Staubli VAL3: insertENDSwitch.pgx

public program insertENDSwitch(string x_sKey, num x_nIndex, bool& x_bToSave)
  local num l_i
begin
  if x_nIndex==0 and progTemp:pProgItem[x_sKey].pProgTemplate[x_nIndex].sTRAJname==""
    x_nIndex=x_nIndex
  else
    x_nIndex=x_nIndex+1
    //// insert(progTemp:pProgItem[x_sKey].pProgTemplate[x_nIndex])
    //l_nIndex=x_nIndex+1
    //insert(progTemp:pProgItem[x_sKey].pProgTemplate[x_nIndex+1])
    append(progTemp:pProgItem[x_sKey].pProgTemplate)
    for l_i = size(progTemp:pProgItem[x_sKey].pProgTemplate)-1 to x_nIndex step -1
      call copyPara(x_sKey,l_i-1,l_i)
    endFor
  endIf

  progTemp:pProgItem[x_sKey].pProgTemplate[x_nIndex].nType=7
  progTemp:pProgItem[x_sKey].pProgTemplate[x_nIndex].sTRAJname="ENDSWITCH"
  x_bToSave=true
end
